(* IEC 61131-3 sources: codesys/project-view/Device/Plc Logic/Application/本机-0-输入输出物理量, 5 files *)

(* ---- GPI.st ---- *)
{attribute 'qualified_only'}
VAR_GLOBAL
	xEStopButton		AT %IX0.0 :BOOL;
	xPauseButton		AT %IX0.1 :BOOL;
	xResetButton		AT %IX0.2 :BOOL;
	xFuntionButton		AT %IX0.3 :BOOL;
	xLocalRackPos1		AT %IX1.4 :BOOL;
	xLocalRackPos2		AT %IX1.5 :BOOL;
	xLocalRackPos3		AT %IX1.6 :BOOL;
	xLocalRackPos4		AT %IX1.7 :BOOL;
END_VAR

(* ---- GPI_Logic.st ---- *)
{attribute 'qualified_only'}
VAR_GLOBAL
	xEStop							:BOOL;
	xPause							:BOOL;
	xContinue						:BOOL;
	xReset							:BOOL;
	xFuntion						:BOOL;
	xLocalRackPos1			AT %MX1000.0:BOOL;
	xLocalRackPos2			AT %MX1002.0:BOOL;
	xLocalRackPos3			AT %MX1004.0:BOOL;
	xLocalRackPos4			AT %MX1006.0:BOOL;
END_VAR

(* ---- GPO.st ---- *)
{attribute 'qualified_only'}
VAR_GLOBAL

END_VAR

(* ---- GPO_Logic.st ---- *)
{attribute 'qualified_only'}
VAR_GLOBAL

END_VAR

(* ---- SR_GPIO.st ---- *)
PROGRAM SR_GPIO
VAR
	rtrigPause					:Standard.R_TRIG;
	ftrigPause					:Standard.F_TRIG;
	rtrigReset					:Standard.R_TRIG;
	rtrigFuntion				:Standard.R_TRIG;
END_VAR
// --- implementation ---
//按钮触发
rtrigPause(CLK:= GPI.xPauseButton, Q=> GPI_Logic.xPause);
ftrigPause(CLK:= GPI.xPauseButton, Q=> GPI_Logic.xContinue);
rtrigReset(CLK:= GPI.xResetButton, Q=> GPI_Logic.xReset);
rtrigFuntion(CLK:= GPI.xFuntionButton, Q=> GPI_Logic.xFuntion);

//传感器滤波处理
GPI_Logic.xLocalRackPos1:=GPI.xLocalRackPos1;
GPI_Logic.xLocalRackPos2:=GPI.xLocalRackPos2;
GPI_Logic.xLocalRackPos3:=GPI.xLocalRackPos3;
GPI_Logic.xLocalRackPos4:=GPI.xLocalRackPos4;
END_PROGRAM
